FUNCTION_BLOCK FB_Valve EXTENDS FB_ValveBase
VAR_OUTPUT
	bOutput	: BOOL;
END_VAR

SUPER^();
bOutput := stStatus.eState = E_ValveState.Open OR stStatus.eState = E_ValveState.Opening;
IF stStatus.eState = E_ValveState.Opening THEN
	stStatus.eState := E_ValveState.Open;
ELSIF stStatus.eState = E_ValveState.Closing THEN
	stStatus.eState := E_ValveState.Closed;
END_IF

ACTION A_Reset:
stStatus.eState := E_ValveState.Closed;
stStatus.nCycles := 0;
bOutput := FALSE;
END_ACTION

METHOD Open : BOOL
VAR_INPUT
	bForce	: BOOL;
END_VAR
Open := SUPER^.Open(bForce := bForce);
IF Open THEN
	bOutput := TRUE;
END_IF
END_METHOD

END_FUNCTION_BLOCK

(* stored: Version 1.1.0.1
   POU FB_Valve: Id {fba7432e-93b5-4bb7-94cd-f1abce3d73ae}, SpecialFunc None
   Action A_Reset: Id {13aabb9b-bde7-4350-aeb5-d561d77ea03b}
   Method Open: Id {02720f70-93be-404c-9c9d-6e37f6846c5f} *)
